PROGRAM ExampleProgram
VAR
END_VAR

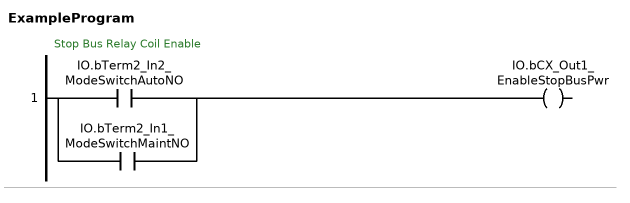
// NETWORK 1
// Stop Bus Relay Coil Enable
IO.bCX_Out1_EnableStopBusPwr := IO.bTerm2_In2_ModeSwitchAutoNO OR IO.bTerm2_In1_ModeSwitchMaintNO;

END_PROGRAM

(* stored: Version 1.1.0.1, ProductVersion 3.1.4024.16
   POU ExampleProgram: Id {ed927ec6-985b-453d-a263-70835cf562cd}, SpecialFunc None *)
